// TIA Portal V21 export
TextList "TL_Order"  ListRange=Decimal
  TextListEntry   Text="0 slobodan redoslijed"
  TextListEntry   From=1, To=1, Text="1 redoslijed po listi"
  TextListEntry   From=2, To=2, Text="2 strogo: istovar pa ukrcaj"
